(*
SPDX-FileCopyrightText: © 2026 Oleksandr Tiutyk <trofimich@gmail.com>
SPDX-License-Identifier: MIT
License: https://opensource.org/license/mit
*)

(*!
<summary>
Beckhoff EP2809_0021: 16-channel digital output EtherCAT Box (24 V DC, 0.5 A, M8).
</summary>
<description>
Process image mapping structure for the EP2809_0021 EtherCAT Box IP67 module with 16 discrete outputs.
When used for I/O, link located fields or their containing buffers to the matching selected PDOs.
The record is not a packed wire buffer; compiler padding is not part of the device specification.
Unlinked/default values do not prove valid I/O. The caller evaluates bus/channel validity before use.
Use one owner task per instance and externally synchronize other access; multi-field snapshots are not atomic.
Copies store data without creating hardware links. Keep borrowed field references valid while consumers are bound.
This passive record performs no validation, synchronization, configuration or protocol advancement.
</description>
*)
TYPE EP2809_0021 :
STRUCT
	Ch01 AT %Q* : BOOL;
	Ch02 AT %Q* : BOOL;
	Ch03 AT %Q* : BOOL;
	Ch04 AT %Q* : BOOL;
	Ch05 AT %Q* : BOOL;
	Ch06 AT %Q* : BOOL;
	Ch07 AT %Q* : BOOL;
	Ch08 AT %Q* : BOOL;
	Ch09 AT %Q* : BOOL;
	Ch10 AT %Q* : BOOL;
	Ch11 AT %Q* : BOOL;
	Ch12 AT %Q* : BOOL;
	Ch13 AT %Q* : BOOL;
	Ch14 AT %Q* : BOOL;
	Ch15 AT %Q* : BOOL;
	Ch16 AT %Q* : BOOL;
END_STRUCT
END_TYPE

(* stored: Version 1.1.0.1, ProductVersion 3.1.4026.20
   DUT EP2809_0021: Id {b45e35f6-87f6-40ff-926f-e4baabecf19d} *)
